(* IEC 61131-3 sources: MongoMation/docs/research/openplc_samples/dialect_tests, 46 files *)

(* ---- t17_user_fb_and_function.st ---- *)
FUNCTION add3 : INT
  VAR_INPUT a : INT; b : INT; c : INT; END_VAR
  add3 := a + b + c;
END_FUNCTION

FUNCTION_BLOCK Latch
  VAR_INPUT set : BOOL; rst : BOOL; END_VAR
  VAR_OUTPUT q : BOOL; END_VAR
  IF rst THEN q := FALSE; ELSIF set THEN q := TRUE; END_IF;
END_FUNCTION_BLOCK

PROGRAM main
  VAR
    l1 : Latch; s : BOOL; r : BOOL; out : BOOL; i : INT;
  END_VAR
  l1(set := s, rst := r);
  out := l1.q;
  i := add3(1, 2, 3);
  i := add3(a := 1, b := 2, c := 3);
END_PROGRAM

CONFIGURATION Config0
  RESOURCE Res0 ON PLC
    TASK task0(INTERVAL := T#20ms,PRIORITY := 0);
    PROGRAM instance0 WITH task0 : main;
  END_RESOURCE
END_CONFIGURATION

(* ---- t44_fb_with_located_inside.st ---- *)
FUNCTION_BLOCK Station
  VAR sensor AT %IX100.0 : BOOL; END_VAR
  VAR_OUTPUT q : BOOL; END_VAR
  q := sensor;
END_FUNCTION_BLOCK
PROGRAM main
  VAR st : Station; y : BOOL; END_VAR
  st();
  y := st.q;
END_PROGRAM

CONFIGURATION Config0
  RESOURCE Res0 ON PLC
    TASK task0(INTERVAL := T#20ms,PRIORITY := 0);
    PROGRAM instance0 WITH task0 : main;
  END_RESOURCE
END_CONFIGURATION

(* ---- t01_line_comment.st ---- *)
PROGRAM main
  VAR
    a : BOOL; // line comment
  END_VAR
  a := NOT a; // toggle
END_PROGRAM

CONFIGURATION Config0
  RESOURCE Res0 ON PLC
    TASK task0(INTERVAL := T#20ms,PRIORITY := 0);
    PROGRAM instance0 WITH task0 : main;
  END_RESOURCE
END_CONFIGURATION

(* ---- t02_block_comment_c_style.st ---- *)
PROGRAM main
  VAR
    a : BOOL; /* C-style block comment */
  END_VAR
  a := NOT a;
END_PROGRAM

CONFIGURATION Config0
  RESOURCE Res0 ON PLC
    TASK task0(INTERVAL := T#20ms,PRIORITY := 0);
    PROGRAM instance0 WITH task0 : main;
  END_RESOURCE
END_CONFIGURATION

(* ---- t03_nested_comment.st ---- *)
PROGRAM main
  VAR
    a : BOOL; (* outer (* inner *) still outer *)
  END_VAR
  a := NOT a;
END_PROGRAM

CONFIGURATION Config0
  RESOURCE Res0 ON PLC
    TASK task0(INTERVAL := T#20ms,PRIORITY := 0);
    PROGRAM instance0 WITH task0 : main;
  END_RESOURCE
END_CONFIGURATION

(* ---- t04_lowercase_keywords.st ---- *)
program main
  var
    a : bool;
    t1 : ton;
  end_var
  t1(in := not a, pt := t#1s);
  if t1.q then a := true; elsif a then a := false; end_if;
end_program

configuration config0
  resource res0 on plc
    task task0(interval := t#20ms, priority := 0);
    program instance0 with task0 : main;
  end_resource
end_configuration

(* ---- t05_no_configuration.st ---- *)
PROGRAM main
  VAR
    a : BOOL;
  END_VAR
  a := NOT a;
END_PROGRAM

(* ---- t06_undeclared_variable.st ---- *)
PROGRAM main
  VAR
    a : BOOL;
  END_VAR
  a := b;
END_PROGRAM

CONFIGURATION Config0
  RESOURCE Res0 ON PLC
    TASK task0(INTERVAL := T#20ms,PRIORITY := 0);
    PROGRAM instance0 WITH task0 : main;
  END_RESOURCE
END_CONFIGURATION

(* ---- t07_type_mismatch_int_to_bool.st ---- *)
PROGRAM main
  VAR
    a : BOOL;
    i : INT := 5;
  END_VAR
  a := i;
END_PROGRAM

CONFIGURATION Config0
  RESOURCE Res0 ON PLC
    TASK task0(INTERVAL := T#20ms,PRIORITY := 0);
    PROGRAM instance0 WITH task0 : main;
  END_RESOURCE
END_CONFIGURATION

(* ---- t08_missing_semicolon.st ---- *)
PROGRAM main
  VAR
    a : BOOL;
  END_VAR
  a := NOT a
END_PROGRAM

CONFIGURATION Config0
  RESOURCE Res0 ON PLC
    TASK task0(INTERVAL := T#20ms,PRIORITY := 0);
    PROGRAM instance0 WITH task0 : main;
  END_RESOURCE
END_CONFIGURATION

(* ---- t09_std_fbs_and_functions.st ---- *)
PROGRAM main
  VAR
    in1 : BOOL; in2 : BOOL; q1 : BOOL; q2 : BOOL; q3 : BOOL; q4 : BOOL; q5 : BOOL; q6 : BOOL;
    i1 : INT := 7; i2 : INT := 3; i3 : INT; r1 : REAL; d1 : DINT; w1 : WORD; t1 : TIME;
    tof1 : TOF; tp1 : TP; ton1 : TON; ft1 : F_TRIG; rt1 : R_TRIG; sr1 : SR; rs1 : RS;
    ctu1 : CTU; ctd1 : CTD; ctud1 : CTUD;
  END_VAR
  tof1(IN := in1, PT := T#2s);
  tp1(IN := in1, PT := T#500ms);
  ton1(IN := in2, PT := TIME#1m30s);
  ft1(CLK := in1);
  rt1(CLK := in2);
  sr1(S1 := in1, R := in2);
  rs1(S := in1, R1 := in2);
  ctu1(CU := rt1.Q, R := ft1.Q, PV := 10);
  ctd1(CD := rt1.Q, LD := ft1.Q, PV := 10);
  ctud1(CU := rt1.Q, CD := ft1.Q, R := FALSE, LD := FALSE, PV := 5);
  q1 := tof1.Q; q2 := tp1.Q; q3 := sr1.Q1; q4 := rs1.Q1; q5 := ctu1.Q; q6 := ctud1.QU;
  i3 := MAX(i1, i2) + MIN(i1, i2) + LIMIT(0, i1, 5) + ABS(-3) + SEL(in1, i1, i2) + MUX(1, i1, i2);
  r1 := INT_TO_REAL(i3) * 1.5 + SQRT(16.0);
  d1 := INT_TO_DINT(i3) * 1000;
  w1 := SHL(INT_TO_WORD(i1), 2) AND 16#FF;
  t1 := ton1.ET + T#100ms;
  IF ton1.ET > T#2s THEN q1 := TRUE; END_IF;
END_PROGRAM

CONFIGURATION Config0
  RESOURCE Res0 ON PLC
    TASK task0(INTERVAL := T#20ms,PRIORITY := 0);
    PROGRAM instance0 WITH task0 : main;
  END_RESOURCE
END_CONFIGURATION

(* ---- t10_write_to_input.st ---- *)
PROGRAM main
  VAR
    sensor AT %IX100.0 : BOOL;
    lamp AT %QX100.0 : BOOL;
  END_VAR
  sensor := TRUE;
  lamp := sensor;
END_PROGRAM

CONFIGURATION Config0
  RESOURCE Res0 ON PLC
    TASK task0(INTERVAL := T#20ms,PRIORITY := 0);
    PROGRAM instance0 WITH task0 : main;
  END_RESOURCE
END_CONFIGURATION

(* ---- t11_global_located_in_config.st ---- *)
PROGRAM main
  VAR_EXTERNAL
    g_sensor : BOOL;
    g_lamp : BOOL;
  END_VAR
  g_lamp := g_sensor;
END_PROGRAM

CONFIGURATION Config0
  VAR_GLOBAL
    g_sensor AT %IX100.0 : BOOL;
    g_lamp AT %QX100.0 : BOOL;
  END_VAR
  RESOURCE Res0 ON PLC
    TASK task0(INTERVAL := T#20ms,PRIORITY := 0);
    PROGRAM instance0 WITH task0 : main;
  END_RESOURCE
END_CONFIGURATION

(* ---- t12_keyword_as_identifier.st ---- *)
PROGRAM main
  VAR
    on : BOOL;
    time : BOOL;
  END_VAR
  on := NOT time;
END_PROGRAM

CONFIGURATION Config0
  RESOURCE Res0 ON PLC
    TASK task0(INTERVAL := T#20ms,PRIORITY := 0);
    PROGRAM instance0 WITH task0 : main;
  END_RESOURCE
END_CONFIGURATION

(* ---- t13_time_literals.st ---- *)
PROGRAM main
  VAR
    t1 : TIME := T#5s; t2 : TIME := TIME#5s; t3 : TIME := t#1m30s; t4 : TIME := T#1.5s; t5 : TIME := T#500MS; t6 : TIME := T#1h2m3s4ms;
  END_VAR
  t1 := t2 + t3;
END_PROGRAM

CONFIGURATION Config0
  RESOURCE Res0 ON PLC
    TASK task0(INTERVAL := T#20ms,PRIORITY := 0);
    PROGRAM instance0 WITH task0 : main;
  END_RESOURCE
END_CONFIGURATION

(* ---- t14_memory_and_word_located.st ---- *)
PROGRAM main
  VAR
    m0 AT %MW0 : INT;
    md0 AT %MD0 : DINT;
    iw AT %IW100 : INT;
    qw AT %QW100 : INT;
    ib AT %IB0 : BYTE;
  END_VAR
  m0 := iw + 1;
  md0 := INT_TO_DINT(m0);
  qw := m0;
END_PROGRAM

CONFIGURATION Config0
  RESOURCE Res0 ON PLC
    TASK task0(INTERVAL := T#20ms,PRIORITY := 0);
    PROGRAM instance0 WITH task0 : main;
  END_RESOURCE
END_CONFIGURATION

(* ---- t15_invalid_bit_index.st ---- *)
PROGRAM main
  VAR
    x AT %IX0.8 : BOOL;
  END_VAR
  VAR
    y : BOOL;
  END_VAR
  y := x;
END_PROGRAM

CONFIGURATION Config0
  RESOURCE Res0 ON PLC
    TASK task0(INTERVAL := T#20ms,PRIORITY := 0);
    PROGRAM instance0 WITH task0 : main;
  END_RESOURCE
END_CONFIGURATION

(* ---- t16_assign_to_constant.st ---- *)
PROGRAM main
  VAR CONSTANT
    K : INT := 5;
  END_VAR
  VAR
    i : INT;
  END_VAR
  K := 6;
  i := K;
END_PROGRAM

CONFIGURATION Config0
  RESOURCE Res0 ON PLC
    TASK task0(INTERVAL := T#20ms,PRIORITY := 0);
    PROGRAM instance0 WITH task0 : main;
  END_RESOURCE
END_CONFIGURATION

(* ---- t18_real_int_mix.st ---- *)
PROGRAM main
  VAR
    r : REAL; i : INT := 3;
  END_VAR
  r := i * 2.5;
END_PROGRAM

CONFIGURATION Config0
  RESOURCE Res0 ON PLC
    TASK task0(INTERVAL := T#20ms,PRIORITY := 0);
    PROGRAM instance0 WITH task0 : main;
  END_RESOURCE
END_CONFIGURATION

(* ---- t19_elseif_keyword.st ---- *)
PROGRAM main
  VAR
    a : BOOL; b : BOOL;
  END_VAR
  IF a THEN b := TRUE; ELSEIF NOT a THEN b := FALSE; END_IF;
END_PROGRAM

CONFIGURATION Config0
  RESOURCE Res0 ON PLC
    TASK task0(INTERVAL := T#20ms,PRIORITY := 0);
    PROGRAM instance0 WITH task0 : main;
  END_RESOURCE
END_CONFIGURATION

(* ---- t20_control_flow_arrays_strings.st ---- *)
PROGRAM main
  VAR
    arr : ARRAY[0..9] OF INT; k : INT; state : INT; s : STRING := 'hello'; n : INT; done : BOOL;
  END_VAR
  FOR k := 0 TO 9 BY 1 DO arr[k] := k * 2; END_FOR;
  WHILE n < 5 DO n := n + 1; END_WHILE;
  REPEAT n := n - 1; UNTIL n <= 0 END_REPEAT;
  CASE state OF
    0: state := 1;
    1, 2: state := 3;
    3..5: done := TRUE; state := 0;
  ELSE state := 0;
  END_CASE;
  s := CONCAT(s, ' world');
  n := LEN(s);
END_PROGRAM

CONFIGURATION Config0
  RESOURCE Res0 ON PLC
    TASK task0(INTERVAL := T#20ms,PRIORITY := 0);
    PROGRAM instance0 WITH task0 : main;
  END_RESOURCE
END_CONFIGURATION

(* ---- t21_positional_fb_call.st ---- *)
PROGRAM main
  VAR
    t1 : TON; a : BOOL;
  END_VAR
  t1(a, T#1s);
END_PROGRAM

CONFIGURATION Config0
  RESOURCE Res0 ON PLC
    TASK task0(INTERVAL := T#20ms,PRIORITY := 0);
    PROGRAM instance0 WITH task0 : main;
  END_RESOURCE
END_CONFIGURATION

(* ---- t22_assign_in_condition.st ---- *)
PROGRAM main
  VAR
    a : BOOL; b : BOOL;
  END_VAR
  IF a := b THEN a := FALSE; END_IF;
END_PROGRAM

CONFIGURATION Config0
  RESOURCE Res0 ON PLC
    TASK task0(INTERVAL := T#20ms,PRIORITY := 0);
    PROGRAM instance0 WITH task0 : main;
  END_RESOURCE
END_CONFIGURATION

(* ---- t23_two_programs_two_tasks.st ---- *)
PROGRAM fast
  VAR a : BOOL; END_VAR
  a := NOT a;
END_PROGRAM
PROGRAM slow
  VAR b : INT; END_VAR
  b := b + 1;
END_PROGRAM
CONFIGURATION Config0
  RESOURCE Res0 ON PLC
    TASK fast_task(INTERVAL := T#10ms,PRIORITY := 0);
    TASK slow_task(INTERVAL := T#100ms,PRIORITY := 1);
    PROGRAM inst_fast WITH fast_task : fast;
    PROGRAM inst_slow WITH slow_task : slow;
  END_RESOURCE
END_CONFIGURATION

(* ---- t24_located_with_initial_value.st ---- *)
PROGRAM main
  VAR
    lamp AT %QX100.0 : BOOL := TRUE;
  END_VAR
  VAR
    x : BOOL;
  END_VAR
  x := lamp;
END_PROGRAM

CONFIGURATION Config0
  RESOURCE Res0 ON PLC
    TASK task0(INTERVAL := T#20ms,PRIORITY := 0);
    PROGRAM instance0 WITH task0 : main;
  END_RESOURCE
END_CONFIGURATION

(* ---- t25_duplicate_location.st ---- *)
PROGRAM main
  VAR
    a AT %QX100.0 : BOOL;
    b AT %QX100.0 : BOOL;
  END_VAR
  a := TRUE; b := FALSE;
END_PROGRAM

CONFIGURATION Config0
  RESOURCE Res0 ON PLC
    TASK task0(INTERVAL := T#20ms,PRIORITY := 0);
    PROGRAM instance0 WITH task0 : main;
  END_RESOURCE
END_CONFIGURATION

(* ---- t26_config_name_not_config0.st ---- *)
PROGRAM main
  VAR a : BOOL; END_VAR
  a := NOT a;
END_PROGRAM
CONFIGURATION MyConfig
  RESOURCE MyRes ON PLC
    TASK task0(INTERVAL := T#20ms,PRIORITY := 0);
    PROGRAM instance0 WITH task0 : main;
  END_RESOURCE
END_CONFIGURATION

(* ---- t27_unused_semicolon_after_end_if_missing.st ---- *)
PROGRAM main
  VAR a : BOOL; b : BOOL; END_VAR
  IF a THEN b := TRUE; END_IF
  a := b;
END_PROGRAM

CONFIGURATION Config0
  RESOURCE Res0 ON PLC
    TASK task0(INTERVAL := T#20ms,PRIORITY := 0);
    PROGRAM instance0 WITH task0 : main;
  END_RESOURCE
END_CONFIGURATION

(* ---- t28_bool_literal_case_and_int_bool_ops.st ---- *)
PROGRAM main
  VAR a : BOOL := True; b : BOOL := false; i : INT; END_VAR
  a := b OR a AND NOT b XOR TRUE;
  i := BOOL_TO_INT(a) + 1;
END_PROGRAM

CONFIGURATION Config0
  RESOURCE Res0 ON PLC
    TASK task0(INTERVAL := T#20ms,PRIORITY := 0);
    PROGRAM instance0 WITH task0 : main;
  END_RESOURCE
END_CONFIGURATION

(* ---- t29_fb_named_like_std_type_conflict.st ---- *)
PROGRAM main
  VAR TON1 : TON; R_TRIG1 : R_TRIG; IN : BOOL; Q : BOOL; END_VAR
  TON1(IN := IN, PT := T#1s);
  Q := TON1.Q;
END_PROGRAM

CONFIGURATION Config0
  RESOURCE Res0 ON PLC
    TASK task0(INTERVAL := T#20ms,PRIORITY := 0);
    PROGRAM instance0 WITH task0 : main;
  END_RESOURCE
END_CONFIGURATION

(* ---- t30_task_without_interval_and_no_with.st ---- *)
PROGRAM main
  VAR a : BOOL; END_VAR
  a := NOT a;
END_PROGRAM
CONFIGURATION Config0
  RESOURCE Res0 ON PLC
    PROGRAM instance0 : main;
  END_RESOURCE
END_CONFIGURATION

(* ---- t31_typed_and_based_literals.st ---- *)
PROGRAM main
  VAR i : INT; w : WORD; b : BYTE; d : DINT; END_VAR
  i := INT#5 + 16#0F + 2#1010 + 8#17;
  w := WORD#16#FFFF;
  b := 16#A5;
  d := DINT#100000;
END_PROGRAM

CONFIGURATION Config0
  RESOURCE Res0 ON PLC
    TASK task0(INTERVAL := T#20ms,PRIORITY := 0);
    PROGRAM instance0 WITH task0 : main;
  END_RESOURCE
END_CONFIGURATION

(* ---- t32_inline_fb_call_in_expression.st ---- *)
PROGRAM main
  VAR rt : R_TRIG; x : BOOL; y : BOOL; END_VAR
  y := rt(CLK := x).Q;
END_PROGRAM

CONFIGURATION Config0
  RESOURCE Res0 ON PLC
    TASK task0(INTERVAL := T#20ms,PRIORITY := 0);
    PROGRAM instance0 WITH task0 : main;
  END_RESOURCE
END_CONFIGURATION

(* ---- t33_bit_access_partial.st ---- *)
PROGRAM main
  VAR w : WORD; x : BOOL; END_VAR
  x := w.0;
END_PROGRAM

CONFIGURATION Config0
  RESOURCE Res0 ON PLC
    TASK task0(INTERVAL := T#20ms,PRIORITY := 0);
    PROGRAM instance0 WITH task0 : main;
  END_RESOURCE
END_CONFIGURATION

(* ---- t34_direct_address_in_code.st ---- *)
PROGRAM main
  VAR x : BOOL; END_VAR
  x := %IX100.0;
  %QX100.0 := x;
END_PROGRAM

CONFIGURATION Config0
  RESOURCE Res0 ON PLC
    TASK task0(INTERVAL := T#20ms,PRIORITY := 0);
    PROGRAM instance0 WITH task0 : main;
  END_RESOURCE
END_CONFIGURATION

(* ---- t35_multi_name_decl.st ---- *)
PROGRAM main
  VAR a, b, c : BOOL; END_VAR
  a := b AND c;
END_PROGRAM

CONFIGURATION Config0
  RESOURCE Res0 ON PLC
    TASK task0(INTERVAL := T#20ms,PRIORITY := 0);
    PROGRAM instance0 WITH task0 : main;
  END_RESOURCE
END_CONFIGURATION

(* ---- t36_int_overflow_literal.st ---- *)
PROGRAM main
  VAR i : INT; END_VAR
  i := 40000;
END_PROGRAM

CONFIGURATION Config0
  RESOURCE Res0 ON PLC
    TASK task0(INTERVAL := T#20ms,PRIORITY := 0);
    PROGRAM instance0 WITH task0 : main;
  END_RESOURCE
END_CONFIGURATION

(* ---- t37_mod_power_exit_return.st ---- *)
PROGRAM main
  VAR i : INT; r : REAL; k : INT; END_VAR
  i := 17 MOD 5;
  r := 2.0 ** 3.0;
  FOR k := 0 TO 10 DO
    IF k = 5 THEN EXIT; END_IF;
  END_FOR;
  IF i = 2 THEN RETURN; END_IF;
  i := i + 1;
END_PROGRAM

CONFIGURATION Config0
  RESOURCE Res0 ON PLC
    TASK task0(INTERVAL := T#20ms,PRIORITY := 0);
    PROGRAM instance0 WITH task0 : main;
  END_RESOURCE
END_CONFIGURATION

(* ---- t38_types_struct_enum.st ---- *)
TYPE
  MotorState : (STOPPED, STARTING, RUNNING, FAULTED);
  Motor : STRUCT
    state : MotorState := STOPPED;
    speed : INT;
  END_STRUCT;
END_TYPE

PROGRAM main
  VAR m : Motor; END_VAR
  CASE m.state OF
    STOPPED: m.state := STARTING;
    STARTING: m.state := RUNNING;
  ELSE m.speed := 0;
  END_CASE;
END_PROGRAM

CONFIGURATION Config0
  RESOURCE Res0 ON PLC
    TASK task0(INTERVAL := T#20ms,PRIORITY := 0);
    PROGRAM instance0 WITH task0 : main;
  END_RESOURCE
END_CONFIGURATION

(* ---- t39_retain_vars.st ---- *)
PROGRAM main
  VAR RETAIN cnt : DINT; END_VAR
  VAR x : BOOL; END_VAR
  cnt := cnt + 1;
END_PROGRAM

CONFIGURATION Config0
  RESOURCE Res0 ON PLC
    TASK task0(INTERVAL := T#20ms,PRIORITY := 0);
    PROGRAM instance0 WITH task0 : main;
  END_RESOURCE
END_CONFIGURATION

(* ---- t40_double_quote_string.st ---- *)
PROGRAM main
  VAR s : STRING; END_VAR
  s := "hello";
END_PROGRAM

CONFIGURATION Config0
  RESOURCE Res0 ON PLC
    TASK task0(INTERVAL := T#20ms,PRIORITY := 0);
    PROGRAM instance0 WITH task0 : main;
  END_RESOURCE
END_CONFIGURATION

(* ---- t41_time_conversions.st ---- *)
PROGRAM main
  VAR t1 : TON; ms : DINT; pt : TIME := T#3s; i : INT; END_VAR
  t1(IN := TRUE, PT := pt);
  ms := TIME_TO_DINT(t1.ET);
  i := DINT_TO_INT(ms / 1000);
  pt := DINT_TO_TIME(5000);
END_PROGRAM

CONFIGURATION Config0
  RESOURCE Res0 ON PLC
    TASK task0(INTERVAL := T#20ms,PRIORITY := 0);
    PROGRAM instance0 WITH task0 : main;
  END_RESOURCE
END_CONFIGURATION

(* ---- t42_empty_statement_and_trailing_comment.st ---- *)
PROGRAM main
  VAR x : BOOL; END_VAR
  ;
  x := NOT x;
END_PROGRAM

CONFIGURATION Config0
  RESOURCE Res0 ON PLC
    TASK task0(INTERVAL := T#20ms,PRIORITY := 0);
    PROGRAM instance0 WITH task0 : main;
  END_RESOURCE
END_CONFIGURATION
(* trailing comment after configuration *)

(* ---- t43_located_in_var_output_of_program.st ---- *)
PROGRAM main
  VAR_OUTPUT lamp AT %QX100.0 : BOOL; END_VAR
  VAR x : BOOL; END_VAR
  lamp := x;
END_PROGRAM

CONFIGURATION Config0
  RESOURCE Res0 ON PLC
    TASK task0(INTERVAL := T#20ms,PRIORITY := 0);
    PROGRAM instance0 WITH task0 : main;
  END_RESOURCE
END_CONFIGURATION

(* ---- t45_real_located_and_int_compare_real.st ---- *)
PROGRAM main
  VAR level AT %IW100 : INT; END_VAR
  VAR pct : REAL; high : BOOL; END_VAR
  pct := INT_TO_REAL(level) / 100.0;
  high := pct > 80;
END_PROGRAM

CONFIGURATION Config0
  RESOURCE Res0 ON PLC
    TASK task0(INTERVAL := T#20ms,PRIORITY := 0);
    PROGRAM instance0 WITH task0 : main;
  END_RESOURCE
END_CONFIGURATION

(* ---- t46_expt_function.st ---- *)
PROGRAM main
  VAR r : REAL; END_VAR
  r := EXPT(2.0, 3.0);
END_PROGRAM

CONFIGURATION Config0
  RESOURCE Res0 ON PLC
    TASK task0(INTERVAL := T#20ms,PRIORITY := 0);
    PROGRAM instance0 WITH task0 : main;
  END_RESOURCE
END_CONFIGURATION
